FUNCTION_BLOCK SolenoidValve IMPLEMENTS I_FillValve, I_Resettable, I_Cyclic
VAR
    _Name          : STRING(32) := 'Solenoid valve';
    _Output        : REFERENCE TO BOOL;
    _OpenFeedback  : REFERENCE TO BOOL;
    _FaultDelay    : TIME;
    _Command       : BOOL;
    _MismatchTimer : TON;
    _IsConfigured  : BOOL;
END_VAR
(*
    SolenoidValve

    Drives one solenoid valve and checks its open-feedback switch. A fault
    is reported while the feedback has disagreed with the command for
    longer than FaultDelay. Name can be set while wiring.
*)

METHOD FB_init : BOOL
VAR_INPUT
    bInitRetains : BOOL;
    bInCopyCode  : BOOL;
    Output       : REFERENCE TO BOOL;
    OpenFeedback : REFERENCE TO BOOL;
    FaultDelay   : TIME;
END_VAR
_Output REF= Output;
_OpenFeedback REF= OpenFeedback;
_FaultDelay := FaultDelay;
_IsConfigured := __ISVALIDREF(Output) AND __ISVALIDREF(OpenFeedback);
END_METHOD

METHOD PUBLIC Open
_Command := TRUE;
END_METHOD

METHOD PUBLIC Close
_Command := FALSE;
END_METHOD

METHOD PUBLIC CyclicLogic
IF NOT _IsConfigured THEN
    RETURN;
END_IF
_Output := _Command;
_MismatchTimer(IN := _Command XOR _OpenFeedback, PT := _FaultDelay);
END_METHOD

METHOD PUBLIC Reset
_MismatchTimer(IN := FALSE);                        // supervise again from now
END_METHOD

PROPERTY PUBLIC IsOpen : BOOL
GET
IsOpen := _IsConfigured AND_THEN (_Command AND _OpenFeedback);
END_GET
END_PROPERTY

PROPERTY PUBLIC IsClosed : BOOL
GET
IsClosed := _IsConfigured AND_THEN NOT (_Command OR _OpenFeedback);
END_GET
END_PROPERTY

PROPERTY PUBLIC HasFault : BOOL
GET
HasFault := NOT _IsConfigured OR _MismatchTimer.Q;
END_GET
END_PROPERTY

PROPERTY PUBLIC FaultText : STRING
GET
IF NOT _IsConfigured THEN
    FaultText := 'I/O not wired';
ELSIF _MismatchTimer.Q THEN
    FaultText := 'No feedback';
ELSE
    FaultText := '';
END_IF
END_GET
END_PROPERTY

PROPERTY PUBLIC Name : STRING
GET
Name := _Name;
END_GET
SET
_Name := Name;
END_SET
END_PROPERTY

END_FUNCTION_BLOCK

(* stored: Version 1.1.0.1, ProductVersion 3.1.4026.0
   POU SolenoidValve: Id {fd880ab6-c8ce-42c9-a59c-218cf7a5749a}, SpecialFunc None
   Folder I_FillValve: Id {4e35492a-8faa-4cee-a833-d6fb69e86dea}
   Folder I_Diagnosable: Id {e5051048-e54b-4183-9fb8-a59ac8df216c}
   Folder I_Resettable: Id {806912db-00f7-4398-b128-85af1f8d730d}
   Folder I_Cyclic: Id {985bb404-9ec5-4ed1-85a8-808c5d994cbf}
   Method FB_init: Id {bb7cce40-1440-4d60-afe9-83ac454f6afd}
   Method Open: Id {7a1466c0-67af-43ea-9e6e-455a9a3b0393}
   Method Close: Id {f35b833f-499e-45c4-a4e1-2cd49cd1bc4d}
   Method CyclicLogic: Id {fd591b0e-e446-4162-bc73-af7e43179407}
   Method Reset: Id {039ab248-d261-4f62-958b-75dd20f668e1}
   Property IsOpen: Id {8371f707-a765-44e8-807f-e43a7d07b20d}
   Get Get: Id {7e5f50db-31f7-4af5-8459-1db6e26d63cf}
   Property IsClosed: Id {6754a114-989f-4e06-81b8-98efc798da79}
   Get Get: Id {100f29e0-7fa5-4fbe-90e5-1ab2ce6d75a9}
   Property HasFault: Id {21d71350-aefb-4f12-b4f1-cd302f40f7ac}
   Get Get: Id {9560971e-e8cf-4fb4-a1c5-3069d47eb8b4}
   Property FaultText: Id {4b72d7cc-454d-4720-8732-d8d84d6fb803}
   Get Get: Id {0b364971-f0fe-404e-b312-a065978fca52}
   Property Name: Id {659692b0-5420-4956-93aa-a22d2e83aaeb}
   Get Get: Id {740a803d-9082-43b5-9cab-6e5c78414479}
   Set Set: Id {865bb9e0-5889-4d66-bb09-92e859702587} *)
